SYSTEM IIOT_AM
  (* Version 1.0, 2020-11-25, eliseu *)
  APPLICATION ARM1
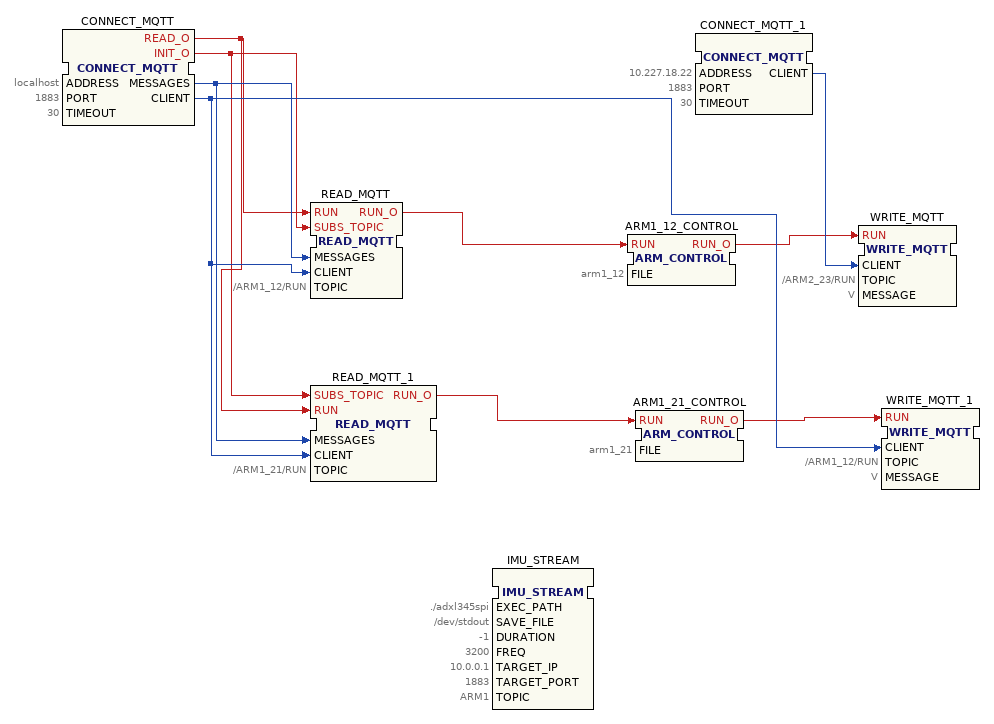
    FBS
      ARM1_12_CONTROL : ARM_CONTROL(FILE := arm1_12);
      ARM1_21_CONTROL : ARM_CONTROL(FILE := arm1_21);
      WRITE_MQTT_1 : WRITE_MQTT(TOPIC := /ARM1_12/RUN, MESSAGE := V);
      READ_MQTT_1 : READ_MQTT(TOPIC := /ARM1_21/RUN);
      WRITE_MQTT : WRITE_MQTT(TOPIC := /ARM2_23/RUN, MESSAGE := V);
      CONNECT_MQTT_1 : CONNECT_MQTT(ADDRESS := 10.227.18.22, PORT := 1883, TIMEOUT := 30);
      CONNECT_MQTT : CONNECT_MQTT(ADDRESS := localhost, PORT := 1883, TIMEOUT := 30);
      READ_MQTT : READ_MQTT(TOPIC := /ARM1_12/RUN);
      IMU_STREAM : IMU_STREAM(EXEC_PATH := ./adxl345spi, SAVE_FILE := /dev/stdout, DURATION := -1, FREQ := 3200, TARGET_IP := 10.0.0.1, TARGET_PORT := 1883, TOPIC := ARM1);
    END_FBS
    EVENT_CONNECTIONS
      CONNECT_MQTT.READ_O TO READ_MQTT.RUN;
      CONNECT_MQTT.INIT_O TO READ_MQTT.SUBS_TOPIC;
      READ_MQTT_1.RUN_O TO ARM1_21_CONTROL.RUN;
      READ_MQTT.RUN_O TO ARM1_12_CONTROL.RUN;
      CONNECT_MQTT.INIT_O TO READ_MQTT_1.SUBS_TOPIC;
      CONNECT_MQTT.READ_O TO READ_MQTT_1.RUN;
      ARM1_12_CONTROL.RUN_O TO WRITE_MQTT.RUN;
      ARM1_21_CONTROL.RUN_O TO WRITE_MQTT_1.RUN;
    END_CONNECTIONS
    DATA_CONNECTIONS
      CONNECT_MQTT_1.CLIENT TO WRITE_MQTT.CLIENT;
      CONNECT_MQTT.MESSAGES TO READ_MQTT.MESSAGES;
      CONNECT_MQTT.MESSAGES TO READ_MQTT_1.MESSAGES;
      CONNECT_MQTT.CLIENT TO READ_MQTT_1.CLIENT;
      CONNECT_MQTT.CLIENT TO WRITE_MQTT_1.CLIENT;
      CONNECT_MQTT.CLIENT TO READ_MQTT.CLIENT;
    END_CONNECTIONS
  END_APPLICATION
  APPLICATION ARM2
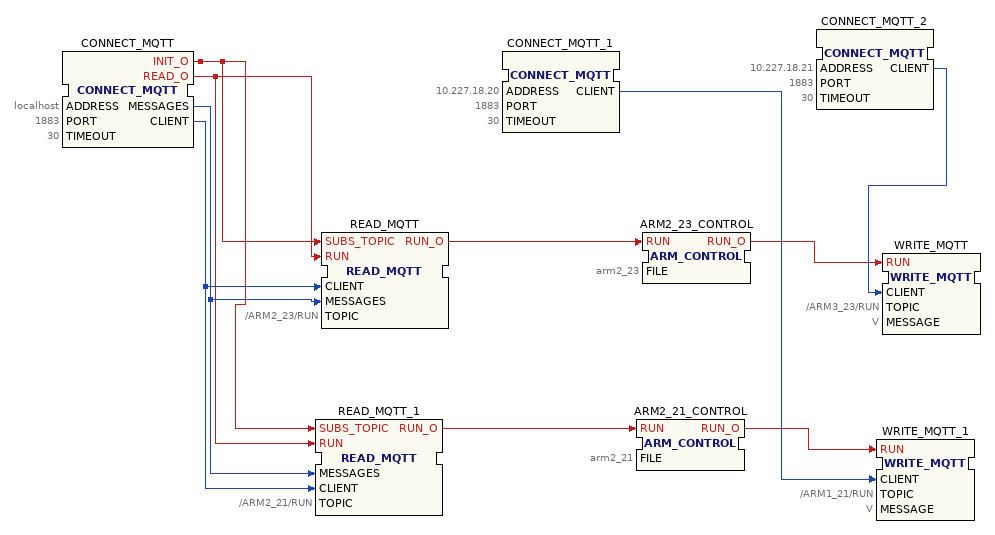
    FBS
      READ_MQTT : READ_MQTT(TOPIC := /ARM2_23/RUN);
      CONNECT_MQTT : CONNECT_MQTT(ADDRESS := localhost, PORT := 1883, TIMEOUT := 30);
      ARM2_21_CONTROL : ARM_CONTROL(FILE := arm2_21);
      WRITE_MQTT : WRITE_MQTT(TOPIC := /ARM3_23/RUN, MESSAGE := V);
      READ_MQTT_1 : READ_MQTT(TOPIC := /ARM2_21/RUN);
      CONNECT_MQTT_2 : CONNECT_MQTT(ADDRESS := 10.227.18.21, PORT := 1883, TIMEOUT := 30);
      ARM2_23_CONTROL : ARM_CONTROL(FILE := arm2_23);
      WRITE_MQTT_1 : WRITE_MQTT(TOPIC := /ARM1_21/RUN, MESSAGE := V);
      CONNECT_MQTT_1 : CONNECT_MQTT(ADDRESS := 10.227.18.20, PORT := 1883, TIMEOUT := 30);
    END_FBS
    EVENT_CONNECTIONS
      READ_MQTT_1.RUN_O TO ARM2_21_CONTROL.RUN;
      CONNECT_MQTT.INIT_O TO READ_MQTT.SUBS_TOPIC;
      ARM2_23_CONTROL.RUN_O TO WRITE_MQTT.RUN;
      CONNECT_MQTT.INIT_O TO READ_MQTT_1.SUBS_TOPIC;
      CONNECT_MQTT.READ_O TO READ_MQTT_1.RUN;
      ARM2_21_CONTROL.RUN_O TO WRITE_MQTT_1.RUN;
      READ_MQTT.RUN_O TO ARM2_23_CONTROL.RUN;
      CONNECT_MQTT.READ_O TO READ_MQTT.RUN;
    END_CONNECTIONS
    DATA_CONNECTIONS
      CONNECT_MQTT.MESSAGES TO READ_MQTT_1.MESSAGES;
      CONNECT_MQTT.CLIENT TO READ_MQTT.CLIENT;
      CONNECT_MQTT_2.CLIENT TO WRITE_MQTT.CLIENT;
      CONNECT_MQTT_1.CLIENT TO WRITE_MQTT_1.CLIENT;
      CONNECT_MQTT.CLIENT TO READ_MQTT_1.CLIENT;
      CONNECT_MQTT.MESSAGES TO READ_MQTT.MESSAGES;
    END_CONNECTIONS
  END_APPLICATION
  APPLICATION ARM3
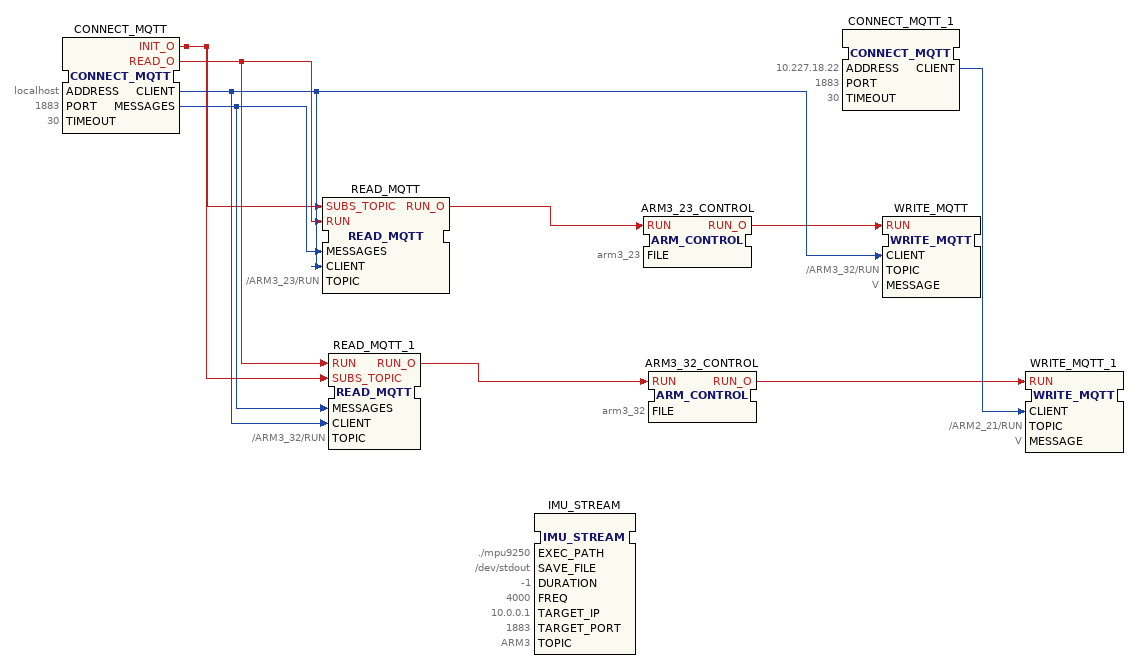
    FBS
      CONNECT_MQTT_1 : CONNECT_MQTT(ADDRESS := 10.227.18.22, PORT := 1883, TIMEOUT := 30);
      CONNECT_MQTT : CONNECT_MQTT(ADDRESS := localhost, PORT := 1883, TIMEOUT := 30);
      ARM3_23_CONTROL : ARM_CONTROL(FILE := arm3_23);
      ARM3_32_CONTROL : ARM_CONTROL(FILE := arm3_32);
      WRITE_MQTT_1 : WRITE_MQTT(TOPIC := /ARM2_21/RUN, MESSAGE := V);
      READ_MQTT_1 : READ_MQTT(TOPIC := /ARM3_32/RUN);
      READ_MQTT : READ_MQTT(TOPIC := /ARM3_23/RUN);
      WRITE_MQTT : WRITE_MQTT(TOPIC := /ARM3_32/RUN, MESSAGE := V);
      IMU_STREAM : IMU_STREAM(EXEC_PATH := ./mpu9250, SAVE_FILE := /dev/stdout, DURATION := -1, FREQ := 4000, TARGET_IP := 10.0.0.1, TARGET_PORT := 1883, TOPIC := ARM3);
    END_FBS
    EVENT_CONNECTIONS
      CONNECT_MQTT.INIT_O TO READ_MQTT.SUBS_TOPIC;
      CONNECT_MQTT.READ_O TO READ_MQTT_1.RUN;
      READ_MQTT.RUN_O TO ARM3_23_CONTROL.RUN;
      CONNECT_MQTT.READ_O TO READ_MQTT.RUN;
      READ_MQTT_1.RUN_O TO ARM3_32_CONTROL.RUN;
      ARM3_32_CONTROL.RUN_O TO WRITE_MQTT_1.RUN;
      ARM3_23_CONTROL.RUN_O TO WRITE_MQTT.RUN;
      CONNECT_MQTT.INIT_O TO READ_MQTT_1.SUBS_TOPIC;
    END_CONNECTIONS
    DATA_CONNECTIONS
      CONNECT_MQTT_1.CLIENT TO WRITE_MQTT_1.CLIENT;
      CONNECT_MQTT.CLIENT TO WRITE_MQTT.CLIENT;
      CONNECT_MQTT.MESSAGES TO READ_MQTT_1.MESSAGES;
      CONNECT_MQTT.MESSAGES TO READ_MQTT.MESSAGES;
      CONNECT_MQTT.CLIENT TO READ_MQTT_1.CLIENT;
      CONNECT_MQTT.CLIENT TO READ_MQTT.CLIENT;
    END_CONNECTIONS
  END_APPLICATION
  APPLICATION PRINTER
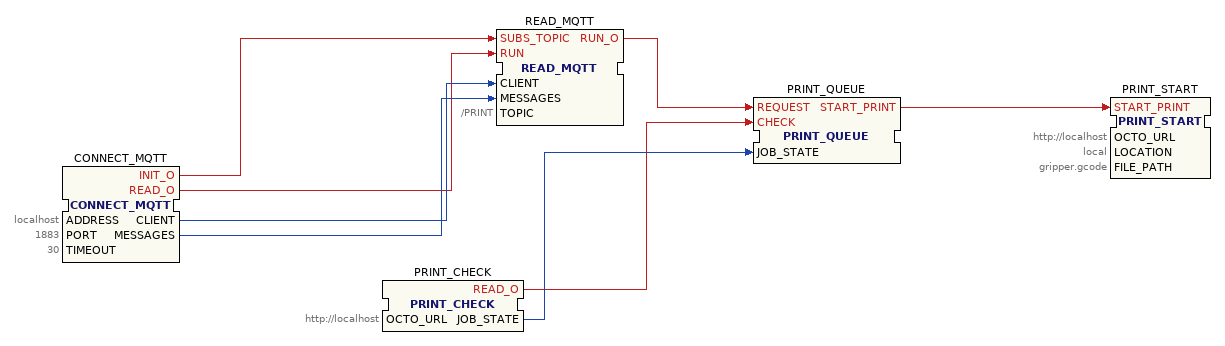
    FBS
      READ_MQTT : READ_MQTT(TOPIC := /PRINT);
      CONNECT_MQTT : CONNECT_MQTT(ADDRESS := localhost, PORT := 1883, TIMEOUT := 30);
      PRINT_CHECK : PRINT_CHECK(OCTO_URL := http://localhost);
      PRINT_QUEUE : PRINT_QUEUE;
      PRINT_START : PRINT_START(OCTO_URL := http://localhost, LOCATION := local, FILE_PATH := gripper.gcode);
    END_FBS
    EVENT_CONNECTIONS
      CONNECT_MQTT.INIT_O TO READ_MQTT.SUBS_TOPIC;
      CONNECT_MQTT.READ_O TO READ_MQTT.RUN;
      READ_MQTT.RUN_O TO PRINT_QUEUE.REQUEST;
      PRINT_QUEUE.START_PRINT TO PRINT_START.START_PRINT;
      PRINT_CHECK.READ_O TO PRINT_QUEUE.CHECK;
    END_CONNECTIONS
    DATA_CONNECTIONS
      CONNECT_MQTT.CLIENT TO READ_MQTT.CLIENT;
      CONNECT_MQTT.MESSAGES TO READ_MQTT.MESSAGES;
      PRINT_CHECK.JOB_STATE TO PRINT_QUEUE.JOB_STATE;
    END_CONNECTIONS
  END_APPLICATION
  APPLICATION PsM1
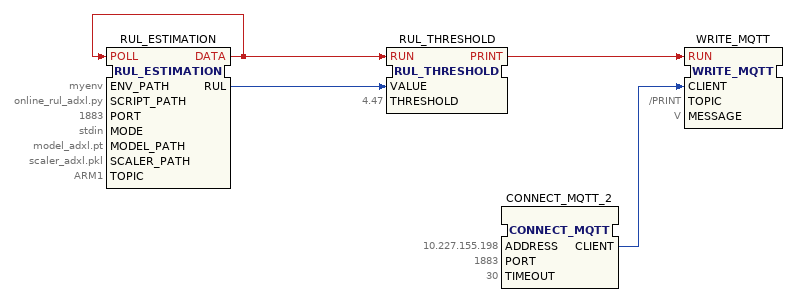
    FBS
      WRITE_MQTT : WRITE_MQTT(TOPIC := /PRINT, MESSAGE := V);
      CONNECT_MQTT_2 : CONNECT_MQTT(ADDRESS := 10.227.155.198, PORT := 1883, TIMEOUT := 30);
      RUL_ESTIMATION : RUL_ESTIMATION(ENV_PATH := myenv, SCRIPT_PATH := online_rul_adxl.py, PORT := 1883, MODE := stdin, MODEL_PATH := model_adxl.pt, SCALER_PATH := scaler_adxl.pkl, TOPIC := ARM1);
      RUL_THRESHOLD : RUL_THRESHOLD(THRESHOLD := 4.47);
    END_FBS
    EVENT_CONNECTIONS
      RUL_ESTIMATION.DATA TO RUL_THRESHOLD.RUN;
      RUL_THRESHOLD.PRINT TO WRITE_MQTT.RUN;
      RUL_ESTIMATION.DATA TO RUL_ESTIMATION.POLL;
    END_CONNECTIONS
    DATA_CONNECTIONS
      CONNECT_MQTT_2.CLIENT TO WRITE_MQTT.CLIENT;
      RUL_ESTIMATION.RUL TO RUL_THRESHOLD.VALUE;
    END_CONNECTIONS
  END_APPLICATION
  APPLICATION PsM2
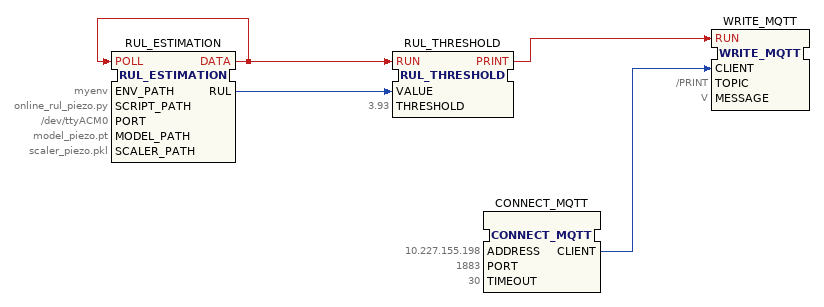
    FBS
      WRITE_MQTT : WRITE_MQTT(TOPIC := /PRINT, MESSAGE := V);
      RUL_THRESHOLD : RUL_THRESHOLD(THRESHOLD := 3.93);
      RUL_ESTIMATION : RUL_ESTIMATION(ENV_PATH := myenv, SCRIPT_PATH := online_rul_piezo.py, PORT := /dev/ttyACM0, MODEL_PATH := model_piezo.pt, SCALER_PATH := scaler_piezo.pkl);
      CONNECT_MQTT : CONNECT_MQTT(ADDRESS := 10.227.155.198, PORT := 1883, TIMEOUT := 30);
    END_FBS
    EVENT_CONNECTIONS
      RUL_ESTIMATION.DATA TO RUL_THRESHOLD.RUN;
      RUL_THRESHOLD.PRINT TO WRITE_MQTT.RUN;
      RUL_ESTIMATION.DATA TO RUL_ESTIMATION.POLL;
    END_CONNECTIONS
    DATA_CONNECTIONS
      RUL_ESTIMATION.RUL TO RUL_THRESHOLD.VALUE;
      CONNECT_MQTT.CLIENT TO WRITE_MQTT.CLIENT;
    END_CONNECTIONS
  END_APPLICATION
  APPLICATION PsM3
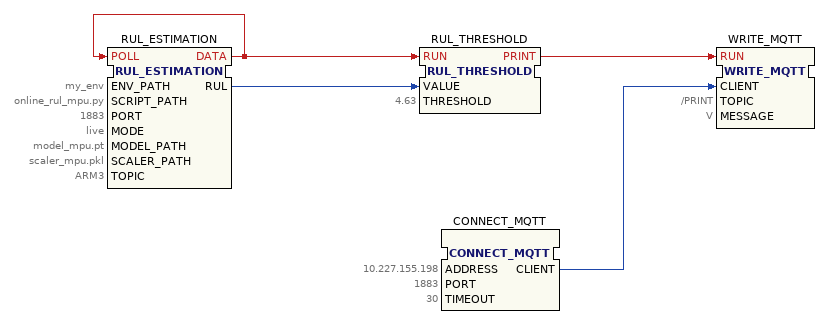
    FBS
      RUL_THRESHOLD : RUL_THRESHOLD(THRESHOLD := 4.63);
      RUL_ESTIMATION : RUL_ESTIMATION(ENV_PATH := my_env, SCRIPT_PATH := online_rul_mpu.py, PORT := 1883, MODE := live, MODEL_PATH := model_mpu.pt, SCALER_PATH := scaler_mpu.pkl, TOPIC := ARM3);
      CONNECT_MQTT : CONNECT_MQTT(ADDRESS := 10.227.155.198, PORT := 1883, TIMEOUT := 30);
      WRITE_MQTT : WRITE_MQTT(TOPIC := /PRINT, MESSAGE := V);
    END_FBS
    EVENT_CONNECTIONS
      RUL_THRESHOLD.PRINT TO WRITE_MQTT.RUN;
      RUL_ESTIMATION.DATA TO RUL_THRESHOLD.RUN;
      RUL_ESTIMATION.DATA TO RUL_ESTIMATION.POLL;
    END_CONNECTIONS
    DATA_CONNECTIONS
      CONNECT_MQTT.CLIENT TO WRITE_MQTT.CLIENT;
      RUL_ESTIMATION.RUL TO RUL_THRESHOLD.VALUE;
    END_CONNECTIONS
  END_APPLICATION
  DEVICE ARM1 : FORTE_PC(MGR_ID := "10.227.18.20:61499")
    {SET_ATTRIBUTE(Profile, HOLOBLOC)} (* device profile *)
    RESOURCE EMB_RES : EMB_RES
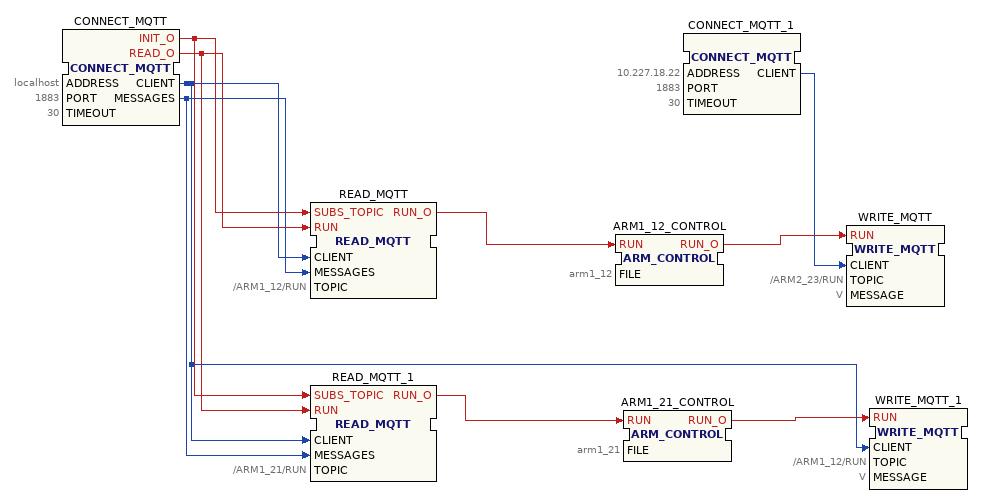
      FBS
        WRITE_MQTT : WRITE_MQTT(TOPIC := /ARM2_23/RUN, MESSAGE := V);
        CONNECT_MQTT : CONNECT_MQTT(ADDRESS := localhost, PORT := 1883, TIMEOUT := 30);
        WRITE_MQTT_1 : WRITE_MQTT(TOPIC := /ARM1_12/RUN, MESSAGE := V);
        READ_MQTT_1 : READ_MQTT(TOPIC := /ARM1_21/RUN);
        ARM1_12_CONTROL : ARM_CONTROL(FILE := arm1_12);
        ARM1_21_CONTROL : ARM_CONTROL(FILE := arm1_21);
        CONNECT_MQTT_1 : CONNECT_MQTT(ADDRESS := 10.227.18.22, PORT := 1883, TIMEOUT := 30);
        READ_MQTT : READ_MQTT(TOPIC := /ARM1_12/RUN);
      END_FBS
      EVENT_CONNECTIONS
        CONNECT_MQTT.INIT_O TO READ_MQTT_1.SUBS_TOPIC;
        CONNECT_MQTT.READ_O TO READ_MQTT_1.RUN;
        READ_MQTT_1.RUN_O TO ARM1_21_CONTROL.RUN;
        CONNECT_MQTT.INIT_O TO READ_MQTT.SUBS_TOPIC;
        CONNECT_MQTT.READ_O TO READ_MQTT.RUN;
        READ_MQTT.RUN_O TO ARM1_12_CONTROL.RUN;
        ARM1_12_CONTROL.RUN_O TO WRITE_MQTT.RUN;
        ARM1_21_CONTROL.RUN_O TO WRITE_MQTT_1.RUN;
      END_CONNECTIONS
      DATA_CONNECTIONS
        CONNECT_MQTT.CLIENT TO WRITE_MQTT_1.CLIENT;
        CONNECT_MQTT.CLIENT TO READ_MQTT_1.CLIENT;
        CONNECT_MQTT.MESSAGES TO READ_MQTT_1.MESSAGES;
        CONNECT_MQTT_1.CLIENT TO WRITE_MQTT.CLIENT;
        CONNECT_MQTT.CLIENT TO READ_MQTT.CLIENT;
        CONNECT_MQTT.MESSAGES TO READ_MQTT.MESSAGES;
      END_CONNECTIONS
    END_RESOURCE
  END_DEVICE
  DEVICE ARM2 : FORTE_PC(MGR_ID := "10.227.18.22:61499")
    {SET_ATTRIBUTE(Profile, HOLOBLOC)} (* device profile *)
    RESOURCE EMB_RES : EMB_RES
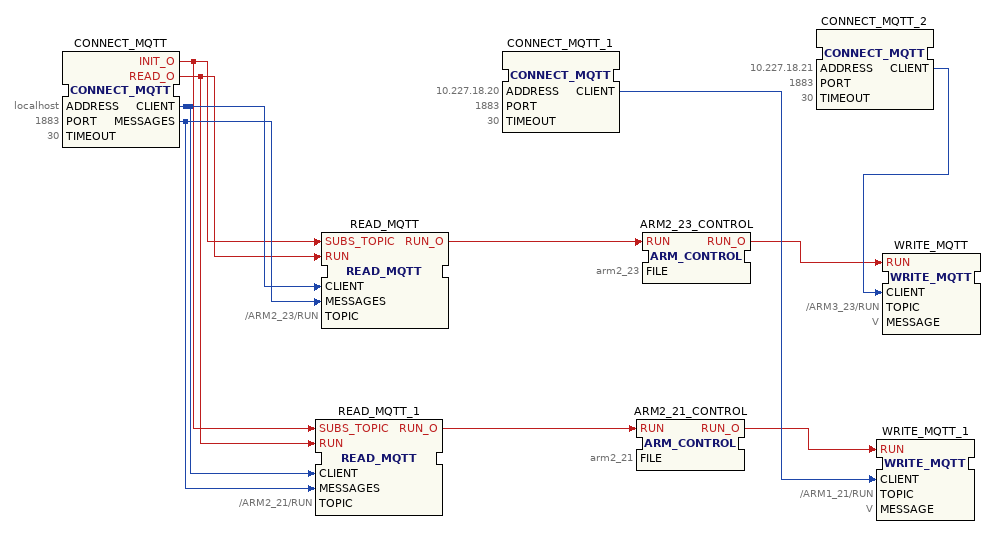
      FBS
        ARM2_23_CONTROL : ARM_CONTROL(FILE := arm2_23);
        READ_MQTT_1 : READ_MQTT(TOPIC := /ARM2_21/RUN);
        WRITE_MQTT_1 : WRITE_MQTT(TOPIC := /ARM1_21/RUN, MESSAGE := V);
        CONNECT_MQTT : CONNECT_MQTT(ADDRESS := localhost, PORT := 1883, TIMEOUT := 30);
        CONNECT_MQTT_2 : CONNECT_MQTT(ADDRESS := 10.227.18.21, PORT := 1883, TIMEOUT := 30);
        READ_MQTT : READ_MQTT(TOPIC := /ARM2_23/RUN);
        WRITE_MQTT : WRITE_MQTT(TOPIC := /ARM3_23/RUN, MESSAGE := V);
        ARM2_21_CONTROL : ARM_CONTROL(FILE := arm2_21);
        CONNECT_MQTT_1 : CONNECT_MQTT(ADDRESS := 10.227.18.20, PORT := 1883, TIMEOUT := 30);
      END_FBS
      EVENT_CONNECTIONS
        CONNECT_MQTT.INIT_O TO READ_MQTT_1.SUBS_TOPIC;
        CONNECT_MQTT.READ_O TO READ_MQTT_1.RUN;
        CONNECT_MQTT.INIT_O TO READ_MQTT.SUBS_TOPIC;
        CONNECT_MQTT.READ_O TO READ_MQTT.RUN;
        READ_MQTT.RUN_O TO ARM2_23_CONTROL.RUN;
        ARM2_23_CONTROL.RUN_O TO WRITE_MQTT.RUN;
        READ_MQTT_1.RUN_O TO ARM2_21_CONTROL.RUN;
        ARM2_21_CONTROL.RUN_O TO WRITE_MQTT_1.RUN;
      END_CONNECTIONS
      DATA_CONNECTIONS
        CONNECT_MQTT.CLIENT TO READ_MQTT_1.CLIENT;
        CONNECT_MQTT.MESSAGES TO READ_MQTT_1.MESSAGES;
        CONNECT_MQTT.CLIENT TO READ_MQTT.CLIENT;
        CONNECT_MQTT.MESSAGES TO READ_MQTT.MESSAGES;
        CONNECT_MQTT_2.CLIENT TO WRITE_MQTT.CLIENT;
        CONNECT_MQTT_1.CLIENT TO WRITE_MQTT_1.CLIENT;
      END_CONNECTIONS
    END_RESOURCE
  END_DEVICE
  DEVICE ARM3 : FORTE_PC(MGR_ID := "10.227.18.21:61499")
    {SET_ATTRIBUTE(Profile, HOLOBLOC)} (* device profile *)
    RESOURCE EMB_RES : EMB_RES
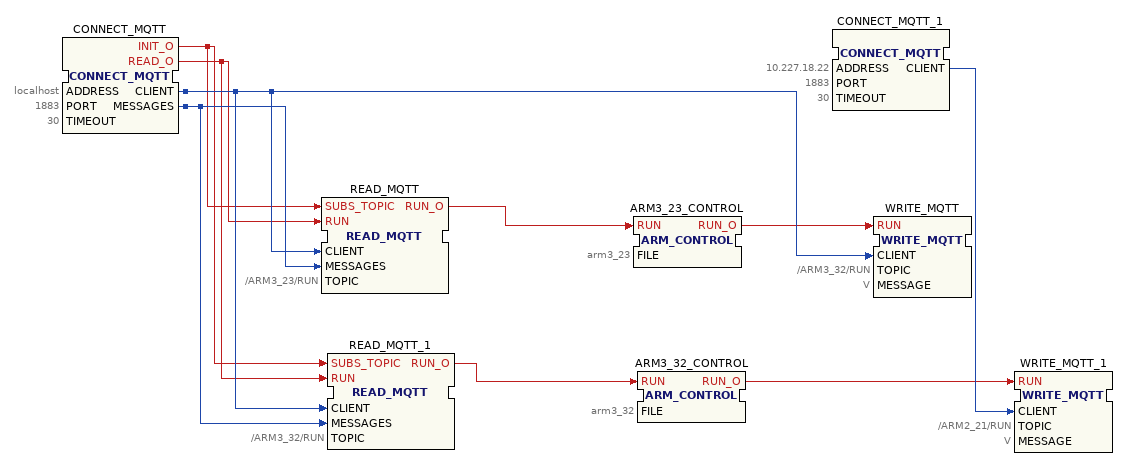
      FBS
        ARM3_32_CONTROL : ARM_CONTROL(FILE := arm3_32);
        WRITE_MQTT_1 : WRITE_MQTT(TOPIC := /ARM2_21/RUN, MESSAGE := V);
        READ_MQTT : READ_MQTT(TOPIC := /ARM3_23/RUN);
        READ_MQTT_1 : READ_MQTT(TOPIC := /ARM3_32/RUN);
        CONNECT_MQTT_1 : CONNECT_MQTT(ADDRESS := 10.227.18.22, PORT := 1883, TIMEOUT := 30);
        WRITE_MQTT : WRITE_MQTT(TOPIC := /ARM3_32/RUN, MESSAGE := V);
        CONNECT_MQTT : CONNECT_MQTT(ADDRESS := localhost, PORT := 1883, TIMEOUT := 30);
        ARM3_23_CONTROL : ARM_CONTROL(FILE := arm3_23);
      END_FBS
      EVENT_CONNECTIONS
        ARM3_32_CONTROL.RUN_O TO WRITE_MQTT_1.RUN;
        READ_MQTT_1.RUN_O TO ARM3_32_CONTROL.RUN;
        CONNECT_MQTT.INIT_O TO READ_MQTT.SUBS_TOPIC;
        CONNECT_MQTT.INIT_O TO READ_MQTT_1.SUBS_TOPIC;
        CONNECT_MQTT.READ_O TO READ_MQTT_1.RUN;
        CONNECT_MQTT.READ_O TO READ_MQTT.RUN;
        READ_MQTT.RUN_O TO ARM3_23_CONTROL.RUN;
        ARM3_23_CONTROL.RUN_O TO WRITE_MQTT.RUN;
      END_CONNECTIONS
      DATA_CONNECTIONS
        CONNECT_MQTT_1.CLIENT TO WRITE_MQTT_1.CLIENT;
        CONNECT_MQTT.CLIENT TO WRITE_MQTT.CLIENT;
        CONNECT_MQTT.CLIENT TO READ_MQTT_1.CLIENT;
        CONNECT_MQTT.CLIENT TO READ_MQTT.CLIENT;
        CONNECT_MQTT.MESSAGES TO READ_MQTT_1.MESSAGES;
        CONNECT_MQTT.MESSAGES TO READ_MQTT.MESSAGES;
      END_CONNECTIONS
    END_RESOURCE
  END_DEVICE
  DEVICE PRINTER : FORTE_PC(MGR_ID := "10.227.155.198:61499")
    {SET_ATTRIBUTE(Profile, HOLOBLOC)} (* device profile *)
    RESOURCE EMB_RES : EMB_RES
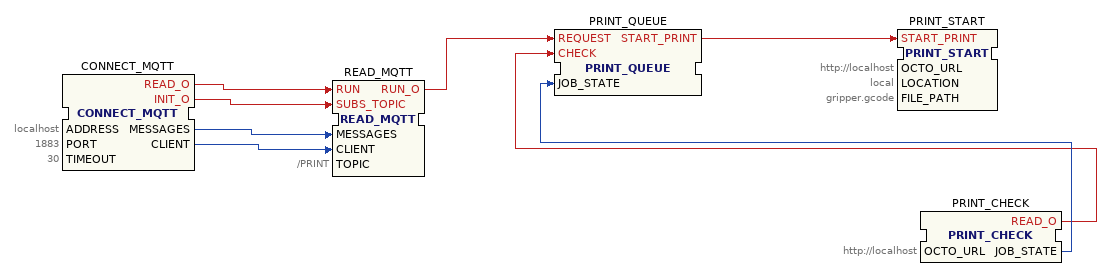
      FBS
        PRINT_START : PRINT_START(OCTO_URL := http://localhost, LOCATION := local, FILE_PATH := gripper.gcode);
        PRINT_QUEUE : PRINT_QUEUE;
        PRINT_CHECK : PRINT_CHECK(OCTO_URL := http://localhost);
        CONNECT_MQTT : CONNECT_MQTT(ADDRESS := localhost, PORT := 1883, TIMEOUT := 30);
        READ_MQTT : READ_MQTT(TOPIC := /PRINT);
      END_FBS
      EVENT_CONNECTIONS
        PRINT_QUEUE.START_PRINT TO PRINT_START.START_PRINT;
        READ_MQTT.RUN_O TO PRINT_QUEUE.REQUEST;
        CONNECT_MQTT.READ_O TO READ_MQTT.RUN;
        CONNECT_MQTT.INIT_O TO READ_MQTT.SUBS_TOPIC;
        PRINT_CHECK.READ_O TO PRINT_QUEUE.CHECK;
      END_CONNECTIONS
      DATA_CONNECTIONS
        PRINT_CHECK.JOB_STATE TO PRINT_QUEUE.JOB_STATE;
        CONNECT_MQTT.MESSAGES TO READ_MQTT.MESSAGES;
        CONNECT_MQTT.CLIENT TO READ_MQTT.CLIENT;
      END_CONNECTIONS
    END_RESOURCE
  END_DEVICE
  DEVICE ARM3_DT : FORTE_PC(MGR_ID := "10.227.18.236:61499")
    {SET_ATTRIBUTE(Profile, HOLOBLOC)} (* device profile *)
    RESOURCE EMB_RES : EMB_RES
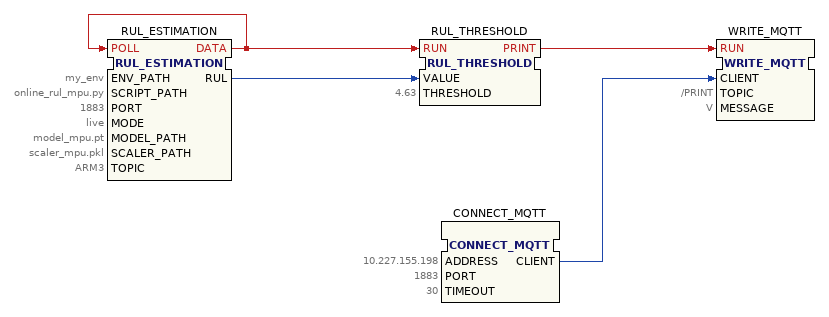
      FBS
        RUL_THRESHOLD : RUL_THRESHOLD(THRESHOLD := 4.63);
        RUL_ESTIMATION : RUL_ESTIMATION(ENV_PATH := my_env, SCRIPT_PATH := online_rul_mpu.py, PORT := 1883, MODE := live, MODEL_PATH := model_mpu.pt, SCALER_PATH := scaler_mpu.pkl, TOPIC := ARM3);
        CONNECT_MQTT : CONNECT_MQTT(ADDRESS := 10.227.155.198, PORT := 1883, TIMEOUT := 30);
        WRITE_MQTT : WRITE_MQTT(TOPIC := /PRINT, MESSAGE := V);
      END_FBS
      EVENT_CONNECTIONS
        RUL_ESTIMATION.DATA TO RUL_ESTIMATION.POLL;
        RUL_ESTIMATION.DATA TO RUL_THRESHOLD.RUN;
        RUL_THRESHOLD.PRINT TO WRITE_MQTT.RUN;
      END_CONNECTIONS
      DATA_CONNECTIONS
        RUL_ESTIMATION.RUL TO RUL_THRESHOLD.VALUE;
        CONNECT_MQTT.CLIENT TO WRITE_MQTT.CLIENT;
      END_CONNECTIONS
    END_RESOURCE
  END_DEVICE
  DEVICE ARM3_SENSOR : FORTE_PC(MGR_ID := "10.227.18.12:61499")
    {SET_ATTRIBUTE(Profile, HOLOBLOC)} (* device profile *)
    RESOURCE EMB_RES : EMB_RES
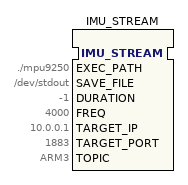
      FBS
        IMU_STREAM : IMU_STREAM(EXEC_PATH := ./mpu9250, SAVE_FILE := /dev/stdout, DURATION := -1, FREQ := 4000, TARGET_IP := 10.0.0.1, TARGET_PORT := 1883, TOPIC := ARM3);
      END_FBS
    END_RESOURCE
  END_DEVICE
  DEVICE ARM2_DT : FORTE_PC(MGR_ID := "10.227.18.211:61499")
    {SET_ATTRIBUTE(Profile, HOLOBLOC)} (* device profile *)
    RESOURCE EMB_RES : EMB_RES
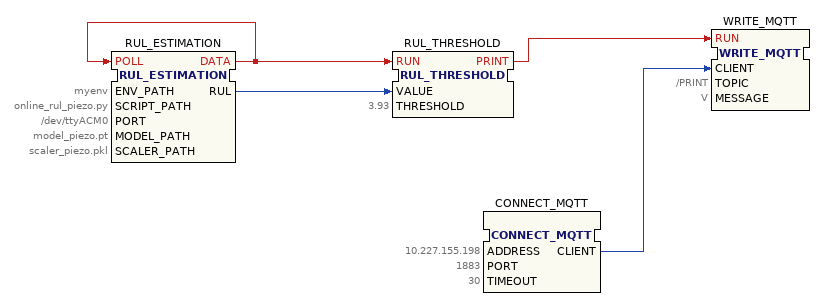
      FBS
        WRITE_MQTT : WRITE_MQTT(TOPIC := /PRINT, MESSAGE := V);
        RUL_THRESHOLD : RUL_THRESHOLD(THRESHOLD := 3.93);
        RUL_ESTIMATION : RUL_ESTIMATION(ENV_PATH := myenv, SCRIPT_PATH := online_rul_piezo.py, PORT := /dev/ttyACM0, MODEL_PATH := model_piezo.pt, SCALER_PATH := scaler_piezo.pkl);
        CONNECT_MQTT : CONNECT_MQTT(ADDRESS := 10.227.155.198, PORT := 1883, TIMEOUT := 30);
      END_FBS
      EVENT_CONNECTIONS
        RUL_THRESHOLD.PRINT TO WRITE_MQTT.RUN;
        RUL_ESTIMATION.DATA TO RUL_ESTIMATION.POLL;
        RUL_ESTIMATION.DATA TO RUL_THRESHOLD.RUN;
      END_CONNECTIONS
      DATA_CONNECTIONS
        RUL_ESTIMATION.RUL TO RUL_THRESHOLD.VALUE;
        CONNECT_MQTT.CLIENT TO WRITE_MQTT.CLIENT;
      END_CONNECTIONS
    END_RESOURCE
  END_DEVICE
  DEVICE ARM1_SENSOR : FORTE_PC(MGR_ID := "10.227.18.15:61499")
    {SET_ATTRIBUTE(Profile, HOLOBLOC)} (* device profile *)
    RESOURCE EMB_RES : EMB_RES
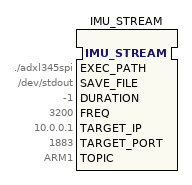
      FBS
        IMU_STREAM : IMU_STREAM(EXEC_PATH := ./adxl345spi, SAVE_FILE := /dev/stdout, DURATION := -1, FREQ := 3200, TARGET_IP := 10.0.0.1, TARGET_PORT := 1883, TOPIC := ARM1);
      END_FBS
    END_RESOURCE
  END_DEVICE
  DEVICE ARM1_DT : FORTE_PC(MGR_ID := "10.227.18.27:61499")
    {SET_ATTRIBUTE(Profile, HOLOBLOC)} (* device profile *)
    RESOURCE EMB_RES : EMB_RES
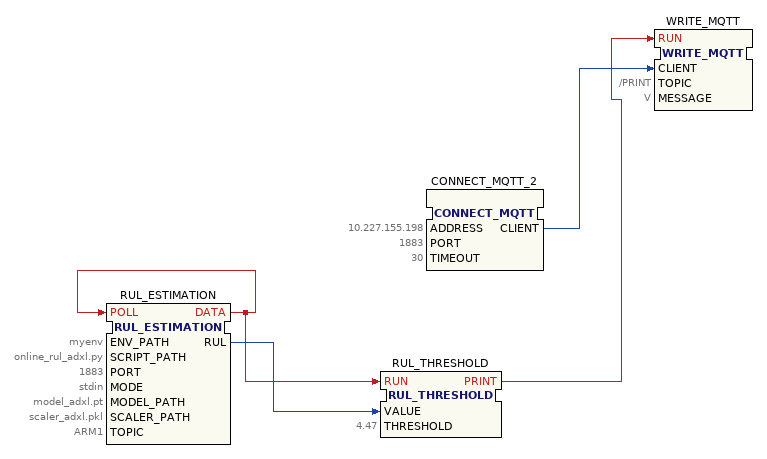
      FBS
        WRITE_MQTT : WRITE_MQTT(TOPIC := /PRINT, MESSAGE := V);
        CONNECT_MQTT_2 : CONNECT_MQTT(ADDRESS := 10.227.155.198, PORT := 1883, TIMEOUT := 30);
        RUL_ESTIMATION : RUL_ESTIMATION(ENV_PATH := myenv, SCRIPT_PATH := online_rul_adxl.py, PORT := 1883, MODE := stdin, MODEL_PATH := model_adxl.pt, SCALER_PATH := scaler_adxl.pkl, TOPIC := ARM1);
        RUL_THRESHOLD : RUL_THRESHOLD(THRESHOLD := 4.47);
      END_FBS
      EVENT_CONNECTIONS
        RUL_ESTIMATION.DATA TO RUL_THRESHOLD.RUN;
        RUL_THRESHOLD.PRINT TO WRITE_MQTT.RUN;
        RUL_ESTIMATION.DATA TO RUL_ESTIMATION.POLL;
      END_CONNECTIONS
      DATA_CONNECTIONS
        CONNECT_MQTT_2.CLIENT TO WRITE_MQTT.CLIENT;
        RUL_ESTIMATION.RUL TO RUL_THRESHOLD.VALUE;
      END_CONNECTIONS
    END_RESOURCE
  END_DEVICE
  MAPPINGS
    ARM1.WRITE_MQTT ON ARM1.EMB_RES.WRITE_MQTT;
    ARM1.CONNECT_MQTT ON ARM1.EMB_RES.CONNECT_MQTT;
    ARM1.WRITE_MQTT_1 ON ARM1.EMB_RES.WRITE_MQTT_1;
    ARM1.READ_MQTT_1 ON ARM1.EMB_RES.READ_MQTT_1;
    ARM1.ARM1_12_CONTROL ON ARM1.EMB_RES.ARM1_12_CONTROL;
    ARM1.ARM1_21_CONTROL ON ARM1.EMB_RES.ARM1_21_CONTROL;
    ARM1.CONNECT_MQTT_1 ON ARM1.EMB_RES.CONNECT_MQTT_1;
    ARM1.READ_MQTT ON ARM1.EMB_RES.READ_MQTT;
    ARM2.ARM2_23_CONTROL ON ARM2.EMB_RES.ARM2_23_CONTROL;
    ARM2.READ_MQTT_1 ON ARM2.EMB_RES.READ_MQTT_1;
    ARM2.WRITE_MQTT_1 ON ARM2.EMB_RES.WRITE_MQTT_1;
    ARM2.CONNECT_MQTT ON ARM2.EMB_RES.CONNECT_MQTT;
    ARM2.CONNECT_MQTT_2 ON ARM2.EMB_RES.CONNECT_MQTT_2;
    ARM2.READ_MQTT ON ARM2.EMB_RES.READ_MQTT;
    ARM2.WRITE_MQTT ON ARM2.EMB_RES.WRITE_MQTT;
    ARM2.ARM2_21_CONTROL ON ARM2.EMB_RES.ARM2_21_CONTROL;
    ARM2.CONNECT_MQTT_1 ON ARM2.EMB_RES.CONNECT_MQTT_1;
    ARM3.ARM3_32_CONTROL ON ARM3.EMB_RES.ARM3_32_CONTROL;
    ARM3.WRITE_MQTT_1 ON ARM3.EMB_RES.WRITE_MQTT_1;
    ARM3.READ_MQTT ON ARM3.EMB_RES.READ_MQTT;
    ARM3.READ_MQTT_1 ON ARM3.EMB_RES.READ_MQTT_1;
    ARM3.CONNECT_MQTT_1 ON ARM3.EMB_RES.CONNECT_MQTT_1;
    ARM3.WRITE_MQTT ON ARM3.EMB_RES.WRITE_MQTT;
    ARM3.CONNECT_MQTT ON ARM3.EMB_RES.CONNECT_MQTT;
    ARM3.ARM3_23_CONTROL ON ARM3.EMB_RES.ARM3_23_CONTROL;
    PsM1.WRITE_MQTT ON ARM1_DT.EMB_RES.WRITE_MQTT;
    PsM1.CONNECT_MQTT_2 ON ARM1_DT.EMB_RES.CONNECT_MQTT_2;
    ARM3.IMU_STREAM ON ARM3_SENSOR.EMB_RES.IMU_STREAM;
    ARM1.IMU_STREAM ON ARM1_SENSOR.EMB_RES.IMU_STREAM;
    PsM1.RUL_ESTIMATION ON ARM1_DT.EMB_RES.RUL_ESTIMATION;
    PsM1.RUL_THRESHOLD ON ARM1_DT.EMB_RES.RUL_THRESHOLD;
    PRINTER.PRINT_START ON PRINTER.EMB_RES.PRINT_START;
    PRINTER.PRINT_QUEUE ON PRINTER.EMB_RES.PRINT_QUEUE;
    PRINTER.PRINT_CHECK ON PRINTER.EMB_RES.PRINT_CHECK;
    PRINTER.CONNECT_MQTT ON PRINTER.EMB_RES.CONNECT_MQTT;
    PRINTER.READ_MQTT ON PRINTER.EMB_RES.READ_MQTT;
    PsM3.RUL_THRESHOLD ON ARM3_DT.EMB_RES.RUL_THRESHOLD;
    PsM3.RUL_ESTIMATION ON ARM3_DT.EMB_RES.RUL_ESTIMATION;
    PsM3.CONNECT_MQTT ON ARM3_DT.EMB_RES.CONNECT_MQTT;
    PsM3.WRITE_MQTT ON ARM3_DT.EMB_RES.WRITE_MQTT;
    PsM2.WRITE_MQTT ON ARM2_DT.EMB_RES.WRITE_MQTT;
    PsM2.RUL_THRESHOLD ON ARM2_DT.EMB_RES.RUL_THRESHOLD;
    PsM2.RUL_ESTIMATION ON ARM2_DT.EMB_RES.RUL_ESTIMATION;
    PsM2.CONNECT_MQTT ON ARM2_DT.EMB_RES.CONNECT_MQTT;
  END_MAPPINGS
  SEGMENTS
    Ethernet : Ethernet;
  END_SEGMENTS
  LINKS
    ARM3 => Ethernet;
    ARM2 => Ethernet;
    ARM1 => Ethernet;
    PRINTER => Ethernet;
    ARM3_DT => Ethernet;
    ARM3_SENSOR => Ethernet;
    ARM2_DT => Ethernet;
    ARM1_SENSOR => Ethernet;
    ARM1_DT => Ethernet;
  END_LINKS
END_SYSTEM
